Fanuc KAREL source: kb00157.KL

-- PROVISIONAL review KL for V770-1; original PC SHA256 d087ddaa93f0174147bd14691080c0c31bb5b0f9556de63b5d656e7d5f397fa2
-- Incomplete behavior may be omitted. Consult companion uncertainty JSON. Do not deploy.
PROGRAM KB00157
%NOLOCKGROUP
BEGIN
  -- UNRESOLVED_PC offsets 5-12; opcodes 9D,23
  -- UNRESOLVED_PC offsets 17-33; opcodes 27,22,31,23
  -- UNRESOLVED_PC offsets 38-42; opcodes 7F
END KB00157
